FUNCTION_BLOCK fbSwitchCtrl
VAR_INPUT
	Switch : iSwitch;
	Config : stSwitchConfig;
END_VAR
VAR_OUTPUT
	State  : stSwitchState;         // Current processed state
    PreviousState  : stSwitchState;         // Previous state
	StateChanged : BOOL;                // State change flag
END_VAR
VAR
	// edge detection
    PressTimerQRise : R_TRIG;
	PressTimerQFall : F_TRIG;
	
    // Timers
    PressTimer : TON;                         // Press duration timer
    MultiClickTimer : TON;                    // Multi-click timer
    
    // Internal
	TempPressCount : USINT := 0;                  // Click counter
	PressTime : TIME := T#0MS;
	ClickType : eSwitchStateType := eSwitchStateType.IDLE;
	
END_VAR
VAR RETAIN
	// Counters
    TotalPresses        : UDINT := 0;          // Total number of clicks
END_VAR

(* 
-----------------------------
fbSwitchController:
Set State output based on Config.Input.
State persist per one PLC cycle, except IDLE, which is a default state.
Every state change sets State.StateChanged to TRUE for one PLC cycle.

SHORT_CLICK <= Config.ShortClickMaxTime
Config.ShortClickMaxTime < LONG_CLICK < Config.LongClickMaxTime
Config.LongClickMaxTime <= HOLD
MULTI_CLICK is multiple SHORT_CLICKs delayed from one another < Config.ShortClickDelayTime
State.PressCount hold amount of switch releases for MULTI_CLICK
-----------------------------
*)

ClickType := eSwitchStateType.IDLE;
StateChanged := FALSE;
PressTimerQRise(CLK := PressTimer.Q);
PressTimerQFall(CLK := PressTimer.Q);

IF Switch.OnPressed THEN
    PressTimer(IN := TRUE, PT := Config.LongClickMaxTime);
END_IF

PressTimer();
MultiClickTimer();

IF Switch.OnReleased THEN
	PressTime := PressTimer.ET;
	PressTimer(IN := FALSE);
	TempPressCount := TempPressCount + 1;
	MultiClickTimer(IN := FALSE);
	
	// Short click
	IF(PressTime <= Config.ShortClickMaxTime) THEN
		MultiClickTimer(IN := TRUE, PT := Config.ShortClickDelayTime);
	// Long click	
	ELSIF (PressTime < Config.LongClickMaxTime) THEN
		ClickType := eSwitchStateType.LONG_CLICK;
	// NOTE: if PressTime = Config.LongClickMaxTime, after HOLD release next state became LONG_CLICK instead of IDLE
	END_IF
END_IF

// Hold click
IF PressTimerQRise.Q THEN
    ClickType := eSwitchStateType.HOLD_ON;
END_IF

IF PressTimerQFall.Q THEN
    ClickType := eSwitchStateType.HOLD_OFF;
END_IF

IF MultiClickTimer.Q THEN
	IF TempPressCount > 1 THEN
		 ClickType := eSwitchStateType.MULTI_CLICK;
	ELSE
		ClickType := eSwitchStateType.SHORT_CLICK;
	END_IF
	MultiClickTimer(IN := FALSE);
END_IF

IF ClickType <> State.StateType THEN
	PreviousState := State;
	State.StateType := ClickType;
	State.PressCount := TempPressCount;
	StateChanged := TRUE;
	TotalPresses     := TotalPresses + 1;
	TempPressCount := 0;
END_IF

END_FUNCTION_BLOCK

(* stored: Version 1.1.0.1
   POU fbSwitchCtrl: Id {d36a5674-47b7-4d99-8111-38bc99505a2d}, SpecialFunc None *)
